(* IEC 61131-3 sources: ZPLC/packages/zplc-ide/plant-scenes/belt-to-sensor, 2 files *)

(* ---- reference.st ---- *)
PROGRAM BeltToSensor
VAR_INPUT
    Start  AT %I0.0 : BOOL;
    EyeFar AT %I0.1 : BOOL;
END_VAR
VAR_OUTPUT
    Run  AT %Q0.0 : BOOL;
    Emit AT %Q0.1 : BOOL;
END_VAR
VAR
    Running : BOOL;
END_VAR

IF Start THEN
    Running := TRUE;
END_IF;
IF EyeFar THEN
    Running := FALSE;
END_IF;

Run := Running;
Emit := Start;

END_PROGRAM

(* ---- starter.st ---- *)
PROGRAM BeltToSensor
VAR_INPUT
    Start  AT %I0.0 : BOOL;  (* StartButton.pressed: the start button *)
    EyeFar AT %I0.1 : BOOL;  (* EyeFar.detect: the sensor at the far end of the belt *)
END_VAR
VAR_OUTPUT
    Run  AT %Q0.0 : BOOL;    (* Belt1.run: run the belt *)
    Emit AT %Q0.1 : BOOL;    (* Emitter1.emit: put one box on the belt *)
END_VAR

(* Goal: a press of the start button puts a box on the belt and runs it;
   the belt stops when the box reaches the far sensor. *)

END_PROGRAM
